Staubli VAL3: SetbtnColor.pgx

public program SetbtnColor(num x_nNum)
  local string l_selColor
  local string l_sNULLcolor
begin
  l_selColor="#9999FF"
  l_sNULLcolor="#FFFFFF"
  switch x_nNum
    case 0
      userPageSet("IO","btn1","style.backgroundColor",l_selColor)
      userPageSet("IO","btn2","style.backgroundColor",l_sNULLcolor)
      userPageSet("IO","btn3","style.backgroundColor",l_sNULLcolor)
      userPageSet("IO","btn4","style.backgroundColor",l_sNULLcolor)
    break
    case 1
      userPageSet("IO","btn1","style.backgroundColor",l_sNULLcolor)
      userPageSet("IO","btn2","style.backgroundColor",l_selColor)
      userPageSet("IO","btn3","style.backgroundColor",l_sNULLcolor)
      userPageSet("IO","btn4","style.backgroundColor",l_sNULLcolor)
    break
    case 2
      userPageSet("IO","btn1","style.backgroundColor",l_sNULLcolor)
      userPageSet("IO","btn2","style.backgroundColor",l_sNULLcolor)
      userPageSet("IO","btn3","style.backgroundColor",l_selColor)
      userPageSet("IO","btn4","style.backgroundColor",l_sNULLcolor)
    break
    case 3
      userPageSet("IO","btn1","style.backgroundColor",l_sNULLcolor)
      userPageSet("IO","btn2","style.backgroundColor",l_sNULLcolor)
      userPageSet("IO","btn3","style.backgroundColor",l_sNULLcolor)
      userPageSet("IO","btn4","style.backgroundColor",l_selColor)
    break
  endSwitch
end
